Fanuc KAREL source: KC00030.KL

PROGRAM KC00030
%NOLOCKGROUP
%ENVIRONMENT UIF
VAR
  I: INTEGER
  J: INTEGER
  K: INTEGER
  R: REAL
  B: BOOLEAN
  S: STRING[80]
  T: STRING[80]
  P: PATH
  Q: PATH
  AI: ARRAY[8] OF INTEGER
  AB: ARRAY[244] OF BYTE
  CD: ARRAY[8] OF COL_DESC_T
  BA: ARRAY[8] OF BOOLEAN
  BC: ARRAY[8,8] OF BOOLEAN
  SA: ARRAY[8] OF STRING[80]
  VP: ARRAY[8,8] OF INTEGER
  X: XWORK_T
BEGIN
  S = 'DICT'
  INIT_TBL(S,I,J,K,CD,BA,BC,SA,VP,X,I)
END KC00030
